Staubli VAL3: Lab2A_Physical.dtx


